// TIA Portal V19 export
FUNCTION_BLOCK "ACT_SPEED_SCALING"   // FB44, LAD
{ S7_Optimized_Access := 'TRUE' }
// stored: AutoNumber false, MemoryReserve 100, SetENOAutomatically false
   VAR_INPUT
      RAW_MIN : Int;
      RAW_MAX : Int;
      SCALE_MIN : Real;
      SCALE_MAX : Real;
      INPUT : Int;
   END_VAR
   VAR_OUTPUT
      SCALE_OUT : Real;
   END_VAR
   VAR
      SP : Real;
   END_VAR
BEGIN

REGION Network 2 (SCL)
   // SPEED SP
   #SP := NORM_X(MIN := #RAW_MIN, VALUE := #INPUT, MAX := #RAW_MIN);
   #SCALE_OUT := SCALE_X(MIN :=#SCALE_MIN, VALUE := #SP, MAX :=#SCALE_MAX);
END_REGION
END_FUNCTION_BLOCK
